KUKA KRL program: LongProg2.src

&ACCESS RVP
&REL 1
&PARAM TEMPLATE = C:\KRC\Roboter\Template\vorgabe
&PARAM EDITMASK = *
DEF LongProg2 ( )
PTP {A1 10.00000,A2 -20.00000,A3 50.00000,A4 0.00000,A5 60.00000,A6 30.00000}
PTP {A1 30.00000,A2 25.00000,A3 80.00000,A4 0.00000,A5 -15.00000,A6 -45.00000}
PTP {A1 10.00000,A2 -20.00000,A3 50.00000,A4 0.00000,A5 60.00000,A6 30.00000}
PTP {A1 30.00000,A2 25.00000,A3 80.00000,A4 0.00000,A5 -15.00000,A6 -45.00000}
PTP {A1 10.00000,A2 -20.00000,A3 50.00000,A4 0.00000,A5 60.00000,A6 30.00000}
END
